Fanuc KAREL source: KC00040.KL

PROGRAM KC00040
%NOLOCKGROUP
%ENVIRONMENT IOSETUP
VAR
  I: INTEGER
  J: INTEGER
  K: INTEGER
  R: REAL
  B: BOOLEAN
  S: STRING[80]
  T: STRING[80]
  P: PATH
  Q: PATH
  AI: ARRAY[8] OF INTEGER
  AB: ARRAY[244] OF BYTE
BEGIN
  GET_PORT_SIM(I,J,B,K)
END KC00040
